screen "AGVs" 1280x800, template "Modèle_1"
   Button "Bouton_3" at 1177,723 size 96x70; TextOff 'IN / OUT'
      on Release: ActivateScreen("Visu_ES-Cpu", 0)
   Button "Bouton_4" at 95,721 size 96x70; TextOff 'Alarmes'
      on Release: ActivateScreen("Alarmes", 0)
      Appearance <- "Bits_B_defaut_en_cours"
   GraphicView "Vue de graphique_5" at 19,728 size 60x60; Picture "Graphique_1"
      Visibility <- "Bits_B_defaut_en_cours"
   Button "Bouton_5" at 1070,723 size 96x70; TextOff 'PARAM'
      on Release: ActivateScreen("Parametrage", 0)
   Button "Bouton_6" at 963,723 size 96x70; TextOff 'MODE MANUEL'
      on Release: ActivateScreen("Mode_Manuel_B01_std_1", 0)
      Appearance <- "Bits_Globaux_x_En_manu"
      ObjectEnable <- "Bits_Globaux_x_En_manu"
   Button "Bouton_7" at 856,723 size 96x70; TextOff 'TP Robots'
      on Click: ActivateScreen("TP_Robots", 0)
      on Release: InvertBit("Bits_B_TP_Robot")
      Appearance <- "B_Pret_TP_Robotique"
   Button "Bouton_8" at 749,723 size 96x70; TextOff 'INIT.'
      on Release: ResetBit("Touche_Tch_Init")
      on Press: SetBit("Touche_Tch_Init")
      Appearance <- "VOY_Init"
      ObjectEnable <- "Bits_Globaux_x_Defaut_non_bloquant"
   Button "Bouton_10" at 535,723 size 96x70; TextOff 'AGVs'
   Button "Bouton_11" at 428,723 size 96x70; TextOff 'Text'
   Button "Bouton_13" at 214,723 size 96x70; TextOff 'Acquit Defaut'
      on Release: ResetBit("Touche_Tch_Acquit")
      on Press: SetBit("Touche_Tch_Acquit")
   Rectangle "Rectangle_15" at 1260,0 size 20x20
      Appearance <- "I_Det_Photo_9"
   Button "Bouton_14" at 4,5 size 124x122; TextOff 'Text'
      on Click: ActivateScreen("Page_demarrage", 0)
   Button "Bouton_9" at 642,723 size 96x70; TextOff 'DEMO. HIPPO'
      on Release: InvertBit("Bits_B_Demo_Hyppo"); ResetBit("Bits_B_TP_Robot")
      Appearance <- "Voyants_HMI_x_VOY_Demo_pret"
      ObjectEnable <- "Bits_Init_glob_OK"
   Button "Bouton_12" at 321,723 size 96x70; TextOff 'HOME'
      on Click: ActivateScreen("Principale", 0)
   Switch "Switch_1" at 270,20 size 120x88; CaptionText 'Changer AGV'; TextOff 'AGV2'; TextOn 'AGV1'
      on SwitchOn: function_efd93a16("AGV2", 8, 133, -1, 2, 1)
      on SwitchOff: function_efd93a16("AGV1", 8, 133, -1, 0, 1)
   Button "Button_1" at 121,216 size 257x136; TextOff 'Lancer boucle GC ABB AMR1'
      on Press: function_b14e0dd5("Touche_Tch_Manu{94}", 0)
   Button "Button_2" at 120,374 size 257x136; TextOff 'Lancer boucle GC UR5 AMR1'
      on Press: function_b14e0dd5("Touche_Tch_Manu{95}", 0)
   Button "Button_3" at 856,215 size 257x136; TextOff 'Lancer boucle PC AMR2'
      on Press: function_b14e0dd5("Touche_Tch_Manu{96}", 0)
*)

(* ===== HMI "HMI_RT_1" =====

ScreenModuleEditorView "Poste Hippodrome" 640x480
   TextField "Champ de texte_34" at 13,13 size 494x21; Text 'Hyppodrome Poste'
   Button "Bouton_1" at 13,64 size 143x58; TextOff 'MONTER BUTEE'
   Button "Bouton_2" at 165,64 size 143x58; TextOff 'DESCENDRE BUTEE'
   Button "Bouton_3" at 13,150 size 143x58; TextOff 'MONTER BUTEE ELEVATEUR'
   Button "Bouton_4" at 165,150 size 143x58; TextOff 'DESCENDRE BUTEE ELEVATEUR'
   Button "Bouton_5" at 13,235 size 143x58; TextOff 'MONTER ELEVATEUR'
   Button "Bouton_6" at 165,235 size 143x58; TextOff 'DESCENDRE ELEVATEUR'
   TextField "Champ de texte_7" at 82,40 size 157x21; Text 'Cmd butée buffer'
   TextField "Champ de texte_8" at 65,125 size 194x21; Text 'Cmd butée elevateur'
   TextField "Champ de texte_9" at 68,210 size 188x21; Text 'Cmd verin elevateur'
   Group "Group" at 315,35 size 202x127
   TextField "Champ de texte_1" at 315,35 size 53x30; Text 'Etat'
   TextField "Champ de texte_2" at 339,62 size 121x23; Text 'Presence pal'
   TextField "Champ de texte_3" at 339,80 size 131x23; Text 'Presence Elev'
   TextField "Champ de texte_4" at 339,99 size 167x23; Text 'Elevateur pos Bas'
   TextField "Champ de texte_5" at 339,118 size 178x23; Text 'Elevateur pos Haut'
   TextField "Champ de texte_10" at 315,139 size 178x23; Text 'Cpt palettes buffer'
   IOField "I/O field_1" at 473,138 size 33x24; FormatPattern 99
   Group "Group_2" at 10,10 size 507x287
   Group "Group_1" at 315,174 size 213x103
   TextField "Champ de texte_6" at 315,174 size 131x30; Text 'Commande'
   TextField "Champ de texte_20" at 336,200 size 134x23; Text 'Rentrer Butée'
   TextField "Champ de texte_21" at 336,218 size 184x23; Text 'Rentrer Butée Elev.'
   TextField "Champ de texte_23" at 336,254 size 192x23; Text 'Descendre Elevateur'
   TextField "Champ de texte_22" at 336,236 size 162x23; Text 'Monter Elevateur'
   Group "Group_3" at 10,10 size 518x287
*)

(* ===== HMI "HMI_RT_1" =====
system functions are stored by id; their names below are inferred from use

ScreenModuleEditorView "Poste Hippodrome" 640x480
   TextField "Champ de texte_34" at 13,13 size 494x21; Text 'Hyppodrome Poste'
   Button "Bouton_1" at 13,64 size 143x58; TextOff 'MONTER BUTEE'
      on Click: ResetBit("DATA_Station.Buffer.cmd.x_Stopper_down")
      Appearance <- "DATA_Station.Buffer.cmd.x_Stopper_down"
   Button "Bouton_2" at 165,64 size 143x58; TextOff 'DESCENDRE BUTEE'
      on Click: SetBit("DATA_Station.Buffer.cmd.x_Stopper_down")
      Appearance <- "DATA_Station.Buffer.cmd.x_Stopper_down"
   Button "Bouton_3" at 13,150 size 143x58; TextOff 'MONTER BUTEE ELEVATEUR'
      on Click: ResetBit("DATA_Station.Elevateur.cmd.x_Stopper_down")
      Appearance <- "DATA_Station.Elevateur.cmd.x_Stopper_down"
   Button "Bouton_4" at 165,150 size 143x58; TextOff 'DESCENDRE BUTEE ELEVATEUR'
      on Click: SetBit("DATA_Station.Elevateur.cmd.x_Stopper_down")
      Appearance <- "DATA_Station.Elevateur.cmd.x_Stopper_down"
   Button "Bouton_5" at 13,235 size 143x58; TextOff 'MONTER ELEVATEUR'
      on Press: function_b14e0dd5("DATA_Station.Elevateur.cmd.x_Elevator_up", 0)
      Appearance <- "DATA_Station.Elevateur.cmd.x_Elevator_up"
   Button "Bouton_6" at 165,235 size 143x58; TextOff 'DESCENDRE ELEVATEUR'
      on Press: function_b14e0dd5("DATA_Station.Elevateur.cmd.x_Elevator_down", 0)
      Appearance <- "DATA_Station.Elevateur.cmd.x_Elevator_down"
   TextField "Champ de texte_7" at 82,40 size 157x21; Text 'Cmd butée buffer'
   TextField "Champ de texte_8" at 65,125 size 194x21; Text 'Cmd butée elevateur'
   TextField "Champ de texte_9" at 68,210 size 188x21; Text 'Cmd verin elevateur'
   TextField "Champ de texte_1" at 315,35 size 53x30; Text 'Etat'
   Rectangle "Rectangle_2" at 317,63 size 17x17
      Appearance <- "DATA_Station.Buffer.status.x_Pres_palette"
   TextField "Champ de texte_2" at 339,62 size 121x23; Text 'Presence pal'
   Rectangle "Rectangle_3" at 317,82 size 17x17
      Appearance <- "DATA_Station.Elevateur.status.x_Pres_palette"
   TextField "Champ de texte_3" at 339,80 size 131x23; Text 'Presence Elev'
   Rectangle "Rectangle_4" at 317,101 size 17x17
      Appearance <- "DATA_Station.Elevateur.status.x_Pos_basse"
   TextField "Champ de texte_4" at 339,99 size 167x23; Text 'Elevateur pos Bas'
   Rectangle "Rectangle_5" at 317,120 size 17x17
      Appearance <- "DATA_Station.Elevateur.status.x_Pos_haute"
   TextField "Champ de texte_5" at 339,118 size 178x23; Text 'Elevateur pos Haut'
   TextField "Champ de texte_6" at 315,174 size 131x30; Text 'Commande'
   Rectangle "Rectangle_23" at 317,202 size 15x16
      Appearance <- "DATA_Station.Buffer.cmd.x_Stopper_down"
   TextField "Champ de texte_20" at 336,200 size 134x23; Text 'Rentrer Butée'
   Rectangle "Rectangle_24" at 317,220 size 15x16
      Appearance <- "DATA_Station.Elevateur.cmd.x_Stopper_down"
   TextField "Champ de texte_21" at 336,218 size 184x23; Text 'Rentrer Butée Elev.'
   Rectangle "Rectangle_25" at 317,238 size 15x16
      Appearance <- "DATA_Station.Elevateur.cmd.x_Elevator_up"
   TextField "Champ de texte_23" at 336,255 size 192x23; Text 'Descendre Elevateur'
   TextField "Champ de texte_22" at 336,237 size 162x23; Text 'Monter Elevateur'
   Rectangle "Rectangle_26" at 317,256 size 15x16
      Appearance <- "DATA_Station.Elevateur.cmd.x_Elevator_down"
   Rectangle "Rectangle_8" at 317,140 size 17x17
      Appearance <- "DATA_Station.Buffer.status.x_buffer_full"
   TextField "Champ de texte_10" at 339,138 size 112x23; Text 'Buffer rempli'
*)

(* ===== HMI "HMI_RT_1" =====
system functions are stored by id; their names below are inferred from use

ScreenModuleEditorView "Poste Hippodrome" 640x480
   TextField "Champ de texte_34" at 13,13 size 494x21; Text 'Hyppodrome Poste'
   Button "Bouton_1" at 13,64 size 143x58; TextOff 'MONTER BUTEE'
      on Click: ResetBit("DATA_Station.Buffer.cmd.x_Stopper_down_manu")
      Appearance <- "DATA_Station.Buffer.cmd.x_Stopper_down_manu"
   Button "Bouton_2" at 165,64 size 143x58; TextOff 'DESCENDRE BUTEE'
      on Click: SetBit("DATA_Station.Buffer.cmd.x_Stopper_down_manu")
      Appearance <- "DATA_Station.Buffer.cmd.x_Stopper_down_manu"
   Button "Bouton_3" at 13,150 size 143x58; TextOff 'MONTER BUTEE ELEVATEUR'
      on Click: ResetBit("DATA_Station.Elevateur.cmd.x_Stopper_down_manual")
      Appearance <- "DATA_Station.Elevateur.cmd.x_Stopper_down_manual"
   Button "Bouton_4" at 165,150 size 143x58; TextOff 'DESCENDRE BUTEE ELEVATEUR'
      on Click: SetBit("DATA_Station.Elevateur.cmd.x_Stopper_down_manual")
      Appearance <- "DATA_Station.Elevateur.cmd.x_Stopper_down_manual"
   Button "Bouton_5" at 13,235 size 143x58; TextOff 'MONTER ELEVATEUR'
      on Press: function_b14e0dd5("DATA_Station.Elevateur.cmd.x_Elevator_up_manual", 0)
      Appearance <- "DATA_Station.Elevateur.cmd.x_Elevator_up_manual"
   Button "Bouton_6" at 165,235 size 143x58; TextOff 'DESCENDRE ELEVATEUR'
      on Press: function_b14e0dd5("DATA_Station.Elevateur.cmd.x_Elevator_down_manual", 0)
      Appearance <- "DATA_Station.Elevateur.cmd.x_Elevator_down_manual"
   TextField "Champ de texte_7" at 82,40 size 157x21; Text 'Cmd butée buffer'
   TextField "Champ de texte_8" at 65,125 size 194x21; Text 'Cmd butée elevateur'
   TextField "Champ de texte_9" at 68,210 size 188x21; Text 'Cmd verin elevateur'
   TextField "Champ de texte_1" at 315,35 size 53x30; Text 'Etat'
   Rectangle "Rectangle_2" at 317,63 size 17x17
      Appearance <- "DATA_Station.Buffer.status.x_Pres_palette"
   TextField "Champ de texte_2" at 339,62 size 121x23; Text 'Presence pal'
   Rectangle "Rectangle_3" at 317,82 size 17x17
      Appearance <- "DATA_Station.Elevateur.status.x_Pres_palette"
   TextField "Champ de texte_3" at 339,80 size 131x23; Text 'Presence Elev'
   Rectangle "Rectangle_4" at 317,101 size 17x17
      Appearance <- "DATA_Station.Elevateur.status.x_Pos_basse"
   TextField "Champ de texte_4" at 339,99 size 167x23; Text 'Elevateur pos Bas'
   Rectangle "Rectangle_5" at 317,120 size 17x17
      Appearance <- "DATA_Station.Elevateur.status.x_Pos_haute"
   TextField "Champ de texte_5" at 339,118 size 178x23; Text 'Elevateur pos Haut'
   TextField "Champ de texte_6" at 315,174 size 131x30; Text 'Commande'
   Rectangle "Rectangle_23" at 317,202 size 15x16
      Appearance <- "DATA_Station.Buffer.cmd.x_Stopper_down"
   TextField "Champ de texte_20" at 336,200 size 134x23; Text 'Rentrer Butée'
   Rectangle "Rectangle_24" at 317,220 size 15x16
      Appearance <- "DATA_Station.Elevateur.cmd.x_Stopper_down"
   TextField "Champ de texte_21" at 336,218 size 184x23; Text 'Rentrer Butée Elev.'
   Rectangle "Rectangle_25" at 317,238 size 15x16
      Appearance <- "DATA_Station.Elevateur.cmd.x_Elevator_up"
   TextField "Champ de texte_23" at 336,255 size 192x23; Text 'Descendre Elevateur'
   TextField "Champ de texte_22" at 336,237 size 162x23; Text 'Monter Elevateur'
   Rectangle "Rectangle_26" at 317,256 size 15x16
      Appearance <- "DATA_Station.Elevateur.cmd.x_Elevator_down"
   Rectangle "Rectangle_8" at 317,140 size 17x17
      Appearance <- "DATA_Station.Buffer.status.x_buffer_full"
   TextField "Champ de texte_10" at 339,138 size 112x23; Text 'Buffer rempli'
*)

(* ===== HMI "HMI_RT_1" =====

ScreenModuleEditorView "Etat_imprimante_3D" 640x480
   TextField "Champ de texte_34" at 136,13 size 140x25; Text 'Imprimante'
   GraphicView "Graphic view_1" at 10,38 size 240x240; Picture "PrusaMK4-noBG"
   TextField "Champ de texte_2" at 254,46 size 63x25; Text 'Ready'
   TextField "Champ de texte_1" at 254,73 size 51x25; Text 'Busy'
   TextField "Champ de texte_3" at 254,103 size 107x25; Text 'Work done'
   TextField "Champ de texte_4" at 254,134 size 99x25; Text 'Home pos'
   TextField "Champ de texte_5" at 254,161 size 127x25; Text 'Print surface'
   TextField "Champ de texte_6" at 254,191 size 53x25; Text 'Fault'
   Button "Button_1" at 227,247 size 168x32; TextOff 'Set workdone'
   TextField "Champ de texte_7" at 254,218 size 153x25; Text 'Work done man'
*)

(* ===== HMI "HMI_RT_1" =====
system functions are stored by id; their names below are inferred from use

ScreenModuleEditorView "Etat_imprimante_3D" 640x480
   TextField "Champ de texte_34" at 136,13 size 140x25; Text 'Imprimante'
   GraphicView "Graphic view_1" at 10,38 size 240x240; Picture "PrusaMK4-noBG"
   Rectangle "Rectangle_2" at 228,49 size 20x20
      Appearance <- "Printer_DATA.Status.x_Ready"
   TextField "Champ de texte_2" at 254,46 size 63x25; Text 'Ready'
   Rectangle "Rectangle_1" at 228,76 size 20x20
      Appearance <- "Printer_DATA.Status.x_Busy"
   TextField "Champ de texte_1" at 254,73 size 51x25; Text 'Busy'
   Rectangle "Rectangle_3" at 228,106 size 20x20
      Appearance <- "Printer_DATA.Status.x_Work_done"
   TextField "Champ de texte_3" at 254,103 size 107x25; Text 'Work done'
   Rectangle "Rectangle_4" at 228,137 size 20x20
      Appearance <- "Printer_DATA.Status.x_AtHome"
   TextField "Champ de texte_4" at 254,134 size 99x25; Text 'Home pos'
   Rectangle "Rectangle_5" at 228,164 size 20x20
      Appearance <- "Printer_DATA.Status.x_HasPrintSurface"
   TextField "Champ de texte_5" at 254,161 size 127x25; Text 'Print surface'
   Rectangle "Rectangle_6" at 228,194 size 20x20
      Appearance <- "Printer_DATA.Status.x_Fault"
   TextField "Champ de texte_6" at 254,191 size 53x25; Text 'Fault'
   Button "Button_1" at 227,247 size 168x32; TextOff 'Set workdone'
      on Press: function_b14e0dd5("Printer_DATA.Status.x_Work_done_manu", 0)
   Rectangle "Rectangle_7" at 228,221 size 20x20
      Appearance <- "Printer_DATA.Status.x_Work_done_manu"
   TextField "Champ de texte_7" at 254,218 size 153x25; Text 'Work done man'
*)

(* ===== HMI "HMI_RT_1" =====
system functions are stored by id; their names below are inferred from use

ScreenModuleEditorView "Poste Hippodrome" 640x480
   TextField "Champ de texte_34" at 13,13 size 494x21; Text 'Hyppodrome Poste'
   Button "Bouton_1" at 13,64 size 143x58; TextOff 'MONTER BUTEE'
      on Click: ResetBit("DATA_Station.Buffer.cmd.x_Stopper_down_manu")
      Appearance <- "DATA_Station.Buffer.cmd.x_Stopper_down_manu"
   Button "Bouton_2" at 165,64 size 143x58; TextOff 'DESCENDRE BUTEE'
      on Click: SetBit("DATA_Station.Buffer.cmd.x_Stopper_down_manu")
      Appearance <- "DATA_Station.Buffer.cmd.x_Stopper_down_manu"
   Button "Bouton_3" at 13,153 size 143x58; TextOff 'MONTER BUTEE ELEVATEUR'
      on Click: ResetBit("DATA_Station.Elevateur.cmd.x_Stopper_down_manual")
      Appearance <- "DATA_Station.Elevateur.cmd.x_Stopper_down_manual"
   Button "Bouton_4" at 165,153 size 143x58; TextOff 'DESCENDRE BUTEE ELEVATEUR'
      on Click: SetBit("DATA_Station.Elevateur.cmd.x_Stopper_down_manual")
      Appearance <- "DATA_Station.Elevateur.cmd.x_Stopper_down_manual"
   Button "Bouton_5" at 13,241 size 143x58; TextOff 'MONTER ELEVATEUR'
      on Press: function_b14e0dd5("DATA_Station.Elevateur.cmd.x_Elevator_up_manual", 0)
      Appearance <- "DATA_Station.Elevateur.cmd.x_Elevator_up_manual"
   Button "Bouton_6" at 165,241 size 143x58; TextOff 'DESCENDRE ELEVATEUR'
      on Press: function_b14e0dd5("DATA_Station.Elevateur.cmd.x_Elevator_down_manual", 0)
      Appearance <- "DATA_Station.Elevateur.cmd.x_Elevator_down_manual"
   TextField "Champ de texte_7" at 82,40 size 157x21; Text 'Cmd butée buffer'
   TextField "Champ de texte_8" at 65,128 size 194x21; Text 'Cmd butée elevateur'
   TextField "Champ de texte_9" at 68,216 size 188x21; Text 'Cmd verin elevateur'
   TextField "Champ de texte_1" at 315,29 size 53x30; Text 'Etat'
   Rectangle "Rectangle_2" at 317,57 size 17x17
      Appearance <- "DATA_Station.Buffer.status.x_Pres_palette"
   TextField "Champ de texte_2" at 339,56 size 121x23; Text 'Presence pal'
   Rectangle "Rectangle_3" at 317,76 size 17x17
      Appearance <- "DATA_Station.Elevateur.status.x_Pres_palette"
   TextField "Champ de texte_3" at 339,74 size 131x23; Text 'Presence Elev'
   Rectangle "Rectangle_4" at 317,95 size 17x17
      Appearance <- "DATA_Station.Elevateur.status.x_Pos_basse"
   TextField "Champ de texte_4" at 339,93 size 167x23; Text 'Elevateur pos Bas'
   Rectangle "Rectangle_5" at 317,114 size 17x17
      Appearance <- "DATA_Station.Elevateur.status.x_Pos_haute"
   TextField "Champ de texte_5" at 339,112 size 178x23; Text 'Elevateur pos Haut'
   TextField "Champ de texte_6" at 315,202 size 131x30; Text 'Commande'
   Rectangle "Rectangle_23" at 317,229 size 15x16
      Appearance <- "DATA_Station.Buffer.cmd.x_Stopper_down"
   TextField "Champ de texte_20" at 336,227 size 134x23; Text 'Rentrer Butée'
   Rectangle "Rectangle_24" at 317,247 size 15x16
      Appearance <- "DATA_Station.Elevateur.cmd.x_Stopper_down"
   TextField "Champ de texte_21" at 336,245 size 184x23; Text 'Rentrer Butée Elev.'
   Rectangle "Rectangle_25" at 317,265 size 15x16
      Appearance <- "DATA_Station.Elevateur.cmd.x_Elevator_up"
   TextField "Champ de texte_23" at 336,282 size 192x23; Text 'Descendre Elevateur'
   TextField "Champ de texte_22" at 336,264 size 162x23; Text 'Monter Elevateur'
   Rectangle "Rectangle_26" at 317,283 size 15x16
      Appearance <- "DATA_Station.Elevateur.cmd.x_Elevator_down"
   Rectangle "Rectangle_8" at 317,133 size 17x17
      Appearance <- "DATA_Station.Buffer.status.x_buffer_full"
   TextField "Champ de texte_10" at 339,131 size 112x23; Text 'Buffer rempli'
   Rectangle "Rectangle_9" at 317,152 size 17x17
      Appearance <- "DATA_Station.Elevateur.status.x_Has_print_surface"
   TextField "Champ de texte_11" at 339,150 size 143x23; Text 'Pres plateau imp'
   Rectangle "Rectangle_10" at 317,171 size 17x17
      Appearance <- "DATA_Station.Elevateur.status.x_Has_3D_piece"
   TextField "Champ de texte_12" at 339,169 size 116x23; Text 'Pres piece 3D'
   Rectangle "Rectangle_11" at 317,190 size 17x17
      Appearance <- "DATA_Station.Elevateur.status.x_Print_surface_clean"
   TextField "Champ de texte_13" at 339,188 size 162x23; Text 'Plateau imp propre'
*)